Fanuc KAREL source: kt00220.KL

PROGRAM KT00220
%STACKSIZE=65535
%PRIORITY=65535
%NOLOCKGROUP
VAR
H1 : ARRAY[2] OF SHORT
I2 : INTEGER
OUT : INTEGER
BEGIN
H1[1]=2
I2=3
-- UNRESOLVED_PC line 10 opcodes [22 9D 33 B3 21 46 23] marker_code=35
END KT00220
